Fanuc KAREL source: kf00103.KL

-- PROVISIONAL review KL for V940-1; original PC SHA256 896c8106534d030267af8b14bb4c4ffdda068d952b70a08bae2462abef8fb382
-- Incomplete behavior may be omitted. Consult companion uncertainty JSON. Do not deploy.
PROGRAM KF00103
%NOLOCKGROUP
BEGIN
  -- V9_ZERO_TABLE_METADATA_HINT layout=0002_ascii; no indexed target words; source/name/runtime held
  -- UNRESOLVED_PC offsets 5-16; opcodes 2E,23
  -- UNRESOLVED_PC offsets 21-32; opcodes 2E,23
  -- UNRESOLVED_PC offsets 37-57; opcodes 27,27,9D,22,2A,22,31
  -- UNRESOLVED_PC offsets 62-66; opcodes 7F
END KF00103
